(* IEC 61131-3 sources: llm-plc-st-eval/codesys/dobles/C3, 7 files *)

(* ---- 01_Correcta.st ---- *)
(* DOBLE DE PRUEBA C3/Correcta - NO ES CORPUS. Esperado: veredicto 1 *)
PROGRAM PRG_Conversion
VAR_INPUT
    btnMarcha : BOOL;
    btnParo : BOOL;
END_VAR
VAR_OUTPUT
    motor : BOOL;
    lampara : BOOL;
END_VAR
VAR
    T1 : TON;
END_VAR
motor := (btnMarcha OR motor) AND NOT btnParo;
T1(IN := motor, PT := T#10S);
lampara := T1.Q;
END_PROGRAM

(* ---- 02_ParoComoNA.st ---- *)
(* DOBLE DE PRUEBA C3/ParoComoNA - NO ES CORPUS. Esperado: veredicto 2, falla en el paso 1 *)
PROGRAM PRG_Conversion
VAR_INPUT
    btnMarcha : BOOL;
    btnParo : BOOL;
END_VAR
VAR_OUTPUT
    motor : BOOL;
    lampara : BOOL;
END_VAR
VAR
    T1 : TON;
END_VAR
motor := (btnMarcha OR motor) AND btnParo;
T1(IN := motor, PT := T#10S);
lampara := T1.Q;
END_PROGRAM

(* ---- 03_SinEnclavamiento.st ---- *)
(* DOBLE DE PRUEBA C3/SinEnclavamiento - NO ES CORPUS. Esperado: veredicto 2, falla en el paso 2 *)
PROGRAM PRG_Conversion
VAR_INPUT
    btnMarcha : BOOL;
    btnParo : BOOL;
END_VAR
VAR_OUTPUT
    motor : BOOL;
    lampara : BOOL;
END_VAR
VAR
    T1 : TON;
END_VAR
motor := btnMarcha AND NOT btnParo;
T1(IN := motor, PT := T#10S);
lampara := T1.Q;
END_PROGRAM

(* ---- 04_MarchaPrioritaria.st ---- *)
(* DOBLE DE PRUEBA C3/MarchaPrioritaria - NO ES CORPUS. Esperado: veredicto 2, falla en el paso 6 *)
PROGRAM PRG_Conversion
VAR_INPUT
    btnMarcha : BOOL;
    btnParo : BOOL;
END_VAR
VAR_OUTPUT
    motor : BOOL;
    lampara : BOOL;
END_VAR
VAR
    T1 : TON;
END_VAR
motor := btnMarcha OR (motor AND NOT btnParo);
T1(IN := motor, PT := T#10S);
lampara := T1.Q;
END_PROGRAM

(* ---- 05_LamparaSinTemporizar.st ---- *)
(* DOBLE DE PRUEBA C3/LamparaSinTemporizar - NO ES CORPUS. Esperado: veredicto 2, falla en el paso 1 *)
PROGRAM PRG_Conversion
VAR_INPUT
    btnMarcha : BOOL;
    btnParo : BOOL;
END_VAR
VAR_OUTPUT
    motor : BOOL;
    lampara : BOOL;
END_VAR
VAR
    T1 : TON;
END_VAR
motor := (btnMarcha OR motor) AND NOT btnParo;
T1(IN := motor, PT := T#10S);
lampara := motor;
END_PROGRAM

(* ---- 06_TiempoCinco.st ---- *)
(* DOBLE DE PRUEBA C3/TiempoCinco - NO ES CORPUS. Esperado: veredicto 2, falla en el paso 2 *)
PROGRAM PRG_Conversion
VAR_INPUT
    btnMarcha : BOOL;
    btnParo : BOOL;
END_VAR
VAR_OUTPUT
    motor : BOOL;
    lampara : BOOL;
END_VAR
VAR
    T1 : TON;
END_VAR
motor := (btnMarcha OR motor) AND NOT btnParo;
T1(IN := motor, PT := T#5S);
lampara := T1.Q;
END_PROGRAM

(* ---- 07_TemporizadorRetenido.st ---- *)
(* DOBLE DE PRUEBA C3/TemporizadorRetenido - NO ES CORPUS. Esperado: veredicto 2, falla en el paso 4 *)
PROGRAM PRG_Conversion
VAR_INPUT
    btnMarcha : BOOL;
    btnParo : BOOL;
END_VAR
VAR_OUTPUT
    motor : BOOL;
    lampara : BOOL;
END_VAR
VAR
    T1 : TON;
END_VAR
motor := (btnMarcha OR motor) AND NOT btnParo;
T1(IN := motor OR T1.Q, PT := T#10S);
lampara := T1.Q;
END_PROGRAM
